FUNCTION_BLOCK AOption_T_2 (* Options-T-Stueck: 1 AOption-Socket IN auf 2 AOption-Plugs OUT1/OUT2 - aktiviert SEQUENZIELL (erst OUT2, nach dessen INIT_CNF erst OUT1), nicht parallel wie AX_SPLIT_2/AR_SPLIT_2. OUT1 kann an den IN-Socket eines weiteren AOption_T_2 angeschlossen werden, um die Kette zu kaskadieren. *)
  (* Standard: 61499-1; Description: Copyright (c) 2026 Meisterschulen am Ostbahnhof This program and the accompanying materials are made available under the terms of the Eclipse Public License 2.0 which is available at https://www.eclipse.org/legal/epl-2.0/ SPDX-License-Identifier: EPL-2.0 *)
  (* Version 1.0, 2026-10-14, Franz Höpfinger, Meisterschulen am Ostbahnhof, initial implementation - generisches, kaskadierbares Gegenstueck zum Ad-hoc-PLUG1-Daisy-Chain-Muster aus OptionalGroup_001a (siehe Uebung_094b3c_AX): statt eine Optionsgruppe selbst um einen Weiterleitungs-Plug zu erweitern, sitzt dieses T-Stueck extern zwischen einem AOption-Ausgang (z.B. eines DEMUX) und beliebig vielen nachgeschalteten Optionsgruppen. Composite statt ECC-BasicFB (Franz) - reines Weiterreichen von Events/QI_OUT, keine eigene Zustandslogik noetig, IEC 61499 Event-Reihenfolge reicht aus. *)
  PACKAGE Option::splitting;
  (* Documentation:
  Sequenzielles T-Stueck fuer AOption
   Nimmt EINEN eingehenden AOption-Request (Socket IN) entgegen und aktiviert daraus ZWEI nachgeschaltete AOption-Verbraucher (Plugs OUT2/OUT1) nacheinander, nicht gleichzeitig: erst OUT2, und erst nachdem dessen INIT_CNF eingetroffen ist, wird OUT1 aktiviert. IN wird erst bestaetigt, wenn BEIDE Ausgaenge bestaetigt haben.
   Deaktivierung laeuft ueber dieselbe Verdrahtung in derselben Reihenfolge (erst OUT2, dann OUT1) - QI_OUT traegt dabei einfach TRUE statt FALSE, die Event-Kette selbst unterscheidet nicht zwischen Aktivierung und Deaktivierung.
   Kaskadierung
   OUT1 kann statt an eine Optionsgruppe an den IN-Socket eines weiteren AOption_T_2 angeschlossen werden - so lassen sich beliebig viele Gruppen streng nacheinander hochfahren, ohne dass eine einzelne Optionsgruppe (wie bisher OptionalGroup_001a) selbst einen Weiterleitungs-Plug mitbringen muss.
   Unterschied zu AX_SPLIT_2/AR_SPLIT_2
   Die bestehenden *_SPLIT_2-Bausteine spiegeln EIN Ereignis/einen Wert PARALLEL auf mehrere Ausgaenge - alle Empfaenger feuern gleichzeitig. Dieses T-Stueck ist bewusst anders: es serialisiert die Aktivierung, damit z.B. eine Gruppe mit Abhaengigkeiten zu einer vorher aktivierten Gruppe sicher erst startet, wenn diese tatsaechlich fertig ist (siehe Uebung_094b3d_AX).
   Warum Composite statt ECC-BasicFB
   Keine eigene Zustandslogik noetig: ein Event feuert erst, wenn sein Quell-Event gefeuert hat - die reine Verkettung IN.INIT_REQ -> OUT2.INIT_REQ -> (wartet auf OUT2.INIT_CNF) -> OUT1.INIT_REQ -> (wartet auf OUT1.INIT_CNF) -> IN.INIT_CNF reicht aus, um dieselbe Sequenzialitaet zu erzwingen wie ein expliziter ECC-Zustandsautomat - ohne InternalVars, ohne Algorithmen.
  *)
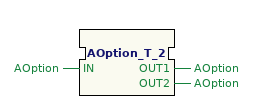
  SOCKETS
    IN : Option::AOption; (* Von einem AOption-Ausgang (z.B. DEMUX.OUTn) gespeist *)
  END_SOCKETS
  PLUGS
    OUT1 : Option::AOption; (* Wird erst nach OUT2.INIT_CNF aktiviert bzw. zuerst deaktiviert - zum Kaskadieren an den IN-Socket eines weiteren AOption_T_2 anschliessbar *)
    OUT2 : Option::AOption; (* Wird zuerst aktiviert (INIT_REQ+) bzw. zuletzt deaktiviert (INIT_REQ-) *)
  END_PLUGS
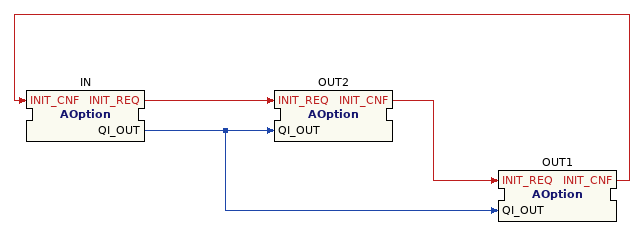
  EVENT_CONNECTIONS
    IN.INIT_REQ TO OUT2.INIT_REQ;
    OUT2.INIT_CNF TO OUT1.INIT_REQ;
    OUT1.INIT_CNF TO IN.INIT_CNF;
  END_CONNECTIONS
  DATA_CONNECTIONS
    IN.QI_OUT TO OUT2.QI_OUT;
    IN.QI_OUT TO OUT1.QI_OUT;
  END_CONNECTIONS
END_FUNCTION_BLOCK
